FUNCTION_BLOCK Distribution (* CAT Function Block Type *)
  (* Standard: 61499-2 *)
  (* Version 0.0, 10/19/2026, Schneider Electric, template *)
  PACKAGE Main;
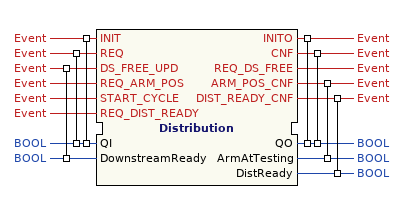
  EVENT_INPUT
    INIT WITH QI; (* Initialization Request *)
    REQ WITH QI; (* Normal Execution Request *)
    DS_FREE_UPD WITH DownstreamReady; (* Update downstream-free state from Testing *)
    REQ_ARM_POS; (* Request current swivel arm-at-Testing status *)
    START_CYCLE; (* Start AutoCycle programmatically *)
    REQ_DIST_READY; (* Request current Distribution ready status *)
  END_EVENT
  EVENT_OUTPUT
    INITO WITH QO; (* Initialization Confirm *)
    CNF WITH QO; (* Execution Confirmation *)
    REQ_DS_FREE; (* Request initial downstream-free status from Testing on startup *)
    ARM_POS_CNF WITH ArmAtTesting; (* Swivel arm-at-Testing status changed *)
    DIST_READY_CNF WITH DistReady; (* Distribution ready state update *)
  END_EVENT
  VAR_INPUT
    QI : BOOL; (* Input event qualifier *)
    DownstreamReady : BOOL; (* Downstream station free state from Testing *)
  END_VAR
  VAR_OUTPUT
    QO : BOOL; (* Output event qualifier *)
    ArmAtTesting : BOOL; (* TRUE when swivel arm is at Testing (3B2) *)
    DistReady : BOOL; (* TRUE when AutoCycle CycleSeq is Stopped or Completed *)
  END_VAR
  FBS
    Ejector : Valve;
    Swivel : Valve2Op;
    Vacuum : Valve;
    BlowOff : DigitalOutput;
    DownstreamFree : DigitalInput;
    MagazineEmpty : DigitalInput;
    EjectorPerm : permCondItem(CondCause := NotActive2, CondName := 'Arm Clear of Magazine', CondPos := Active1);
    Reset : ResetSequence;
    Cycle : AutoCycle;
    DsConv : ANY2ANY_143E21D40326C8151; {SET_ATTRIBUTE(Configuration.GenericFBType.InterfaceParams, Runtime.Standard#CNT:=1;IN${CNT$}:BOOL;OUT${CNT$}:VTQBOOL)}
    DsLink : SYMLINKMULTIVARSRC_298DC1F529059FB5(QI := TRUE, NAME1 := 'RES0.Distribution.DownstreamFree.pv.DIn'); {SET_ATTRIBUTE(Configuration.GenericFBType.InterfaceParams, Runtime.System#I:=1;VALUE${I$}:VTQBOOL)}
    ArmPosOut : AND_550FE6D62F509EB3(IN2 := TRUE, IN3 := TRUE); {SET_ATTRIBUTE(Configuration.GenericFBType.InterfaceParams, Runtime.Standard#CNT:=3;OUT:BOOL)}
    NotDistStop : NOT_42C76073DCEB1A7A; {SET_ATTRIBUTE(Configuration.GenericFBType.InterfaceParams, Runtime.Standard#CNT:=1;OUT${CNT$}:BOOL)}
    NotDistComp : NOT_42C76073DCEB1A7A; {SET_ATTRIBUTE(Configuration.GenericFBType.InterfaceParams, Runtime.Standard#CNT:=1;OUT${CNT$}:BOOL)}
    DistBusyAnd : AND_550FE6D62F509EB3(IN3 := TRUE); {SET_ATTRIBUTE(Configuration.GenericFBType.InterfaceParams, Runtime.Standard#CNT:=3;OUT:BOOL)}
    DistReadyOut : NOT_42C76073DCEB1A7A; {SET_ATTRIBUTE(Configuration.GenericFBType.InterfaceParams, Runtime.Standard#CNT:=1;OUT${CNT$}:BOOL)}
  END_FBS
  EVENT_CONNECTIONS
    Vacuum.CNF TO Reset.FECC89DB3D2A57FF;
    Swivel.CNF TO Reset.A5069DC6B641011A;
    Ejector.CNF TO Reset.43498683653FD650;
    INIT TO Reset.9D471DE3BB9549E0;
    INIT TO Cycle.A729492442D0C9A1;
    Vacuum.CNF TO Cycle.5D63E5C8B975CEB9;
    Swivel.CNF TO Cycle.2CDF47D3663E6E3F;
    Ejector.CNF TO Cycle.FB025A14BE6C5638;
    MagazineEmpty.CNF TO Cycle.7119241BD2443AA1;
    DownstreamFree.CNF TO Cycle.6490AF8BD623FEB6;
    INIT TO DsLink.INIT;
    DsLink.INITO TO REQ_DS_FREE;
    DsLink.INITO TO DsConv.REQ;
    DS_FREE_UPD TO DsConv.REQ;
    DsConv.CNF TO DsLink.REQ;
    INIT TO ArmPosOut.REQ;
    REQ_ARM_POS TO ArmPosOut.REQ;
    Swivel.CNF TO ArmPosOut.REQ;
    ArmPosOut.CNF TO ARM_POS_CNF;
    START_CYCLE TO Cycle.A1B2000000000001;
    INIT TO NotDistStop.REQ;
    REQ_DIST_READY TO NotDistStop.REQ;
    Cycle.A1B2000000000002 TO NotDistStop.REQ;
    NotDistStop.CNF TO NotDistComp.REQ;
    NotDistComp.CNF TO DistBusyAnd.REQ;
    DistBusyAnd.CNF TO DistReadyOut.REQ;
    DistReadyOut.CNF TO DIST_READY_CNF;
  END_CONNECTIONS
  DATA_CONNECTIONS
    Vacuum.FbClosed TO Reset.60387A5202353395;
    Swivel.FbClosed TO Reset.DDDAB227DF90F2E9;
    Ejector.FbClosed TO Reset.22FAB5CD31E08CC4;
    Vacuum.FbOpened TO Cycle.102E354520A9B5EF;
    Vacuum.FbClosed TO Cycle.3E0D46D015AC4734;
    Ejector.FbClosed TO Cycle.F50145A9F34B3204;
    Ejector.FbOpened TO Cycle.27E5B1CA69BBB159;
    Swivel.FbClosed TO Cycle.038D0D4E12791418;
    Swivel.FbOpen TO Cycle.279E4466CE606266;
    Swivel.FbStopped TO Reset.7A3C1E904B2D8F15;
    Swivel.FbStopped TO Cycle.9F1C4E72A38D6B05;
    MagazineEmpty.Pv TO Cycle.795155DF007843B9;
    DownstreamFree.Pv TO Cycle.041FFAAD79F17532;
    DownstreamReady TO DsConv.IN1;
    DsConv.OUT1 TO DsLink.VALUE1;
    Swivel.FbOpen TO ArmPosOut.IN1;
    ArmPosOut.OUT TO ArmAtTesting;
    Cycle.A1B2000000000003 TO NotDistStop.IN1;
    Cycle.A1B2000000000004 TO NotDistComp.IN1;
    NotDistStop.OUT1 TO DistBusyAnd.IN1;
    NotDistComp.OUT1 TO DistBusyAnd.IN2;
    DistBusyAnd.OUT TO DistReadyOut.IN1;
    DistReadyOut.OUT1 TO DistReady;
  END_CONNECTIONS
  ADAPTER_CONNECTIONS
    Swivel.IFbState TO EjectorPerm.ICondSignal;
    EjectorPerm.ICondChainOut TO Ejector.IPerm;
  END_CONNECTIONS
END_FUNCTION_BLOCK
